// TIA Portal V21 export
// export: Created 2026-08-21T20:18:50.8741333Z, ExportSetting None, DisplayName Totally Integrated Automation Portal, DisplayVersion V21, DisplayName STEP 7 Professional, DisplayVersion V21, DisplayName STEP 7 Safety, DisplayVersion V21, DisplayName Tech WebApplication, DisplayVersion V21, DisplayName WinCC Basic/Comfort/Advanced, DisplayVersion V21, DisplayName WinCC Professional, DisplayVersion V21, DisplayName WinCC Unified, DisplayVersion V21
FUNCTION "LAH100" : Void   // FC8, FBD
{ S7_Optimized_Access := 'TRUE' }
// stored: SetENOAutomatically false
BEGIN

REGION Network 1: MonDiL
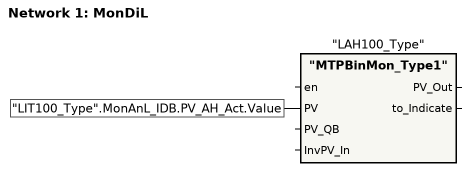
   "LAH100_Type"(PV := "LIT100_Type".MonAnL_IDB.PV_AH_Act.Value);   // "MTPBinMon_Type1"
END_REGION
END_FUNCTION
